Universal Robots URScript: hello_world.script

# HEADER_BEGIN

def test_func():
  textmsg("test function")
  popup("Hello external control", blocking = True)
end

# HEADER_END

# NODE_CONTROL_LOOP_BEGINS

test_func()

# NODE_CONTROL_LOOP_ENDS
